// TIA Portal V21 export
// export: Created 2026-11-08T21:35:25.5370827Z, ExportSetting WithDefaults, DisplayName Totally Integrated Automation Portal, DisplayVersion V21 Update 3, DisplayName STEP 7 Professional, DisplayVersion V21 Update 3, DisplayName STEP 7 Safety, DisplayVersion V21, DisplayName Tech WebApplication, DisplayVersion V21, DisplayName WinCC Basic/Comfort/Advanced, DisplayVersion V21 Update 3, DisplayName WinCC Unified, DisplayVersion V21 Update 3
FUNCTION_BLOCK "FB_StlC_021"   // FB91, STL
TITLE = STL call NE_TypeOfDB
{ S7_Optimized_Access := 'TRUE' }
VERSION : 0.1
// stored: AutoNumber true, IsRetainMemResEnabled false, MemoryReserve 100, UDAEnableTagReadback false
   VAR_INPUT
      dba : DB_ANY;
   END_VAR
   VAR_OUTPUT
      "b" : Bool;
   END_VAR
BEGIN

NETWORK
TITLE = 021 NE_TypeOfDB
      CALL  NE_TypeOfDB
      ( IN1     := #dba,
        IN2     := IEC_TIMER,
        Ret_Val := #"b"
      );
END_FUNCTION_BLOCK
